// TwinCAT 3 PLC project TrsClientTester
// ProgramVersion: 3.1.4023.0
// libraries:
//   ESO LDC Timer Library, * (ESO)
//   Tc2_EtherCAT, * (Beckhoff Automation GmbH)
//   Tc2_Standard, * (Beckhoff Automation GmbH)
//   Tc2_System, * (Beckhoff Automation GmbH)
//   Tc2_Utilities, * (Beckhoff Automation GmbH)
//   Tc3_Module, * (Beckhoff Automation GmbH)
//   VisuDialogs, * (System)
// project tree:
//   DUTs/Enumerations/ E_TEST_STATE.TcDUT
//   / GlobalTextList.TcGTLO, PlcTask.TcTTO, Visualization Manager.TcVMO (not stored)
//   POUs/ MAIN.TcPOU
//   VISUs/ GUI_TIME.TcVIS, GUI_TIMER.TcVIS
// real-time tasks:
//   TASK PlcTask: cycle T#1ms, priority 20, ADS port 350
// I/O:
//   DEVICE Device 1 (EtherCAT), AmsNetId 198.19.191.40.2.1
//     Term 1 (EK1200) [EK1200-5000 EtherCAT Power supply (2A E-Bus)]
//       Term 2 (EK1110) [EK1110 EtherCAT extension]
//     Term 3 (EK1100) [EK1100 EtherCAT Coupler (2A E-Bus)]
//       Term 4 (EL2262) [EL2262 2Ch. Dig. Output 24V, 1µs, DC Oversample]
//       Term 5 (EL6688) [EL6688 - External Synchronisation Interface (IEEE1588)]
//       Term 6 (EL9011) [EL9011 End Terminal]
//   DEVICE Device 5 (NOV-DP-RAM)
//   DEVICE Device 2 (RT-Ethernet Adapter)
// variable links:
//   TrsClientTester/TrsClientTester Instance <-> Device 1 (EtherCAT)
//     PlcTask Inputs/MAIN.fbTimeObj.i_dc2ExtOffset <-> InfoData/DcToExtTimeOffset
//     PlcTask Inputs/MAIN.fbTimeObj.i_dc2TcOffset <-> InfoData/DcToTcTimeOffset
//   TrsClientTester/TrsClientTester Instance <-> Device 1 (EtherCAT)/Term 3 (EK1100)/Term 4 (EL2262)
//     PlcTask Inputs/MAIN.fbTimerObj.DcOutputShift <-> InfoData/DcOutputShift
//     PlcTask Outputs/MAIN.fbTimerObj.CyclicCounter <-> CycCount0/Cycle Counter0
//     PlcTask Outputs/MAIN.fbTimerObj.Output0[{1..125}] <-> Sample0 {0..124}/Output0  (125 links)
//   TrsClientTester/TrsClientTester Instance <-> Device 1 (EtherCAT)/Term 3 (EK1100)/Term 5 (EL6688)
//     PlcTask Inputs/MAIN.fbTimeObj.i_AdsAddr <-> InfoData/AdsAddr
//     PlcTask Inputs/MAIN.fbTimeObj.i_exTime <->   External Sync/External time stamp
//     PlcTask Inputs/MAIN.fbTimeObj.i_extDevNotConnected <->   External Sync/External device not connected
//     PlcTask Inputs/MAIN.fbTimeObj.i_inTime <->   External Sync/Internal time stamp

CONFIGURATION TrsClientTester
    RESOURCE PLC ON TwinCAT3
        TASK PlcTask(INTERVAL := T#1ms, PRIORITY := 20);
        PROGRAM MAIN WITH PlcTask : MAIN;
    END_RESOURCE
END_CONFIGURATION

// ---- DUTs/Enumerations/E_TEST_STATE.TcDUT
{attribute 'qualified_only'}
{attribute 'strict'}
TYPE E_TEST_STATE :
(
	STATE_TEST_OFF				:= 0,
	STATE_TEST_RUNNING
);
END_TYPE

// ---- POUs/MAIN.TcPOU
PROGRAM MAIN
VAR
	fbTimeObj: FB_TIME;
	fbTimerObj: FB_TIMER;
	
	
END_VAR

fbTimeObj();

fbTimerObj(fbTimerRef := fbTimeObj);

END_PROGRAM

// ---- VISUs/GUI_TIME.TcVIS
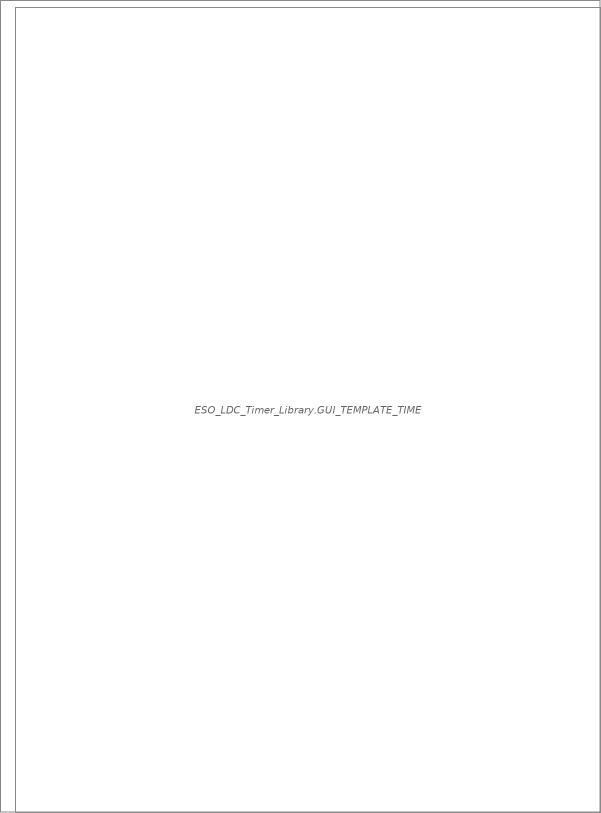
VISUALIZATION GUI_TIME  // 601x813
    Frame (15,7 586x806)
        shows ESO_LDC_Timer_Library.GUI_TEMPLATE_TIME(m_DeviceName := 'timer', m_Instance := MAIN.fbTimeObj)
END_VISUALIZATION

// ---- VISUs/GUI_TIMER.TcVIS
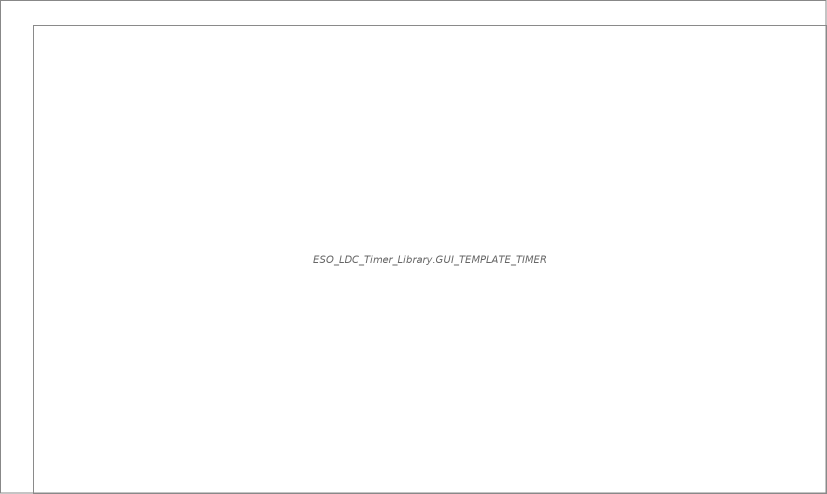
VISUALIZATION GUI_TIMER  // 827x494
    Frame (33,25 794x469)
        shows ESO_LDC_Timer_Library.GUI_TEMPLATE_TIMER(m_Instance := MAIN.fbTimerObj)
END_VISUALIZATION
